INTERFACE ITcoSequencer EXTENDS ITcoState

(*~
	<docu>
		<summary>
			Gets the information about the current step.						
		</summary>				
	</docu>	
~*)
PROPERTY CurrentStep : REFERENCE TO StepDetails
GET
END_GET
END_PROPERTY

PROPERTY ModeController : ITcoSequencerModeController
GET
END_GET
END_PROPERTY

(*~
	<docu>
		<summary>
			<para>
				Ensures calling the Open(), Main() and Close() methods in the desired order.
				This method is final, so it cannot be overloaded. The InstanceName.Run() needs to be called cyclically inside the appropriate context.
			</para>
		</summary>			
	</docu>	
~*)
METHOD PUBLIC FINAL Run
END_METHOD

END_INTERFACE

(* stored: Version 1.1.0.1
   Itf ITcoSequencer: Id {a8c5aaea-ce66-4699-94d6-6fc2b0db7583}
   Property CurrentStep: Id {9693bfe8-b533-07e4-0b7f-afb04386f3c0}
   Get Get: Id {d55c7f61-ec4e-07a2-2f32-e75c01fe1a25}
   Property ModeController: Id {dd9b56ed-8b06-0f8b-10a4-bc7f86421e90}
   Get Get: Id {c118fb9b-2261-0bb2-3940-3e2e9974072b}
   Method Run: Id {c085653a-ddfd-0ace-0d80-e733121bd868} *)
